Fanuc KAREL source: KO00034.KL

PROGRAM KO00034
%NOLOCKGROUP
%ENVIRONMENT MIR
VAR
  P1: POSITION
  P2: POSITION
  F: BOOLEAN
  OUT: XYZWPR
BEGIN
  F = TRUE
  OUT = MIRROR(P1, P2, F)
END KO00034
